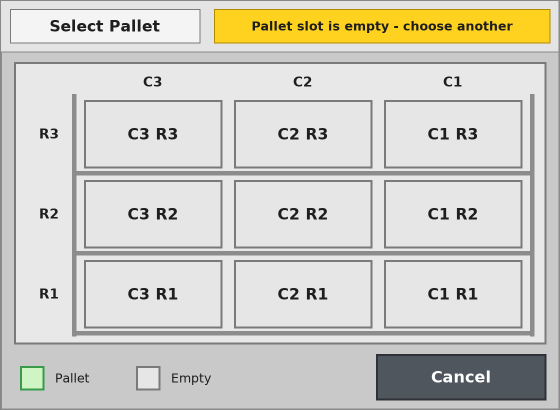
VISUALIZATION SelectPalletDialog  // 560x410
    Rectangle (0,0 560x410)
    Rectangle (0,0 560x52)
    Rectangle (10,9 190x34), "Select Pallet"
    Rectangle (214,12 334x28), "Tap a green slot to retrieve the pallet"
    RoundedRectangle (14,62 532x282)
    Rectangle (84,70 138x24), "C3"
    Rectangle (234,70 138x24), "C2"
    Rectangle (384,70 138x24), "C1"
    Rectangle (24,100 50x68), "R3"
    Rectangle (24,180 50x68), "R2"
    Rectangle (24,260 50x68), "R1"
    Rectangle (72,94 4x242)
    Rectangle (530,94 4x242)
    Rectangle (72,171 462x4)
    Rectangle (72,251 462x4)
    Rectangle (72,331 462x4)
    RoundedRectangle (84,100 138x68), "C3 R3", colour toggle: MAIN.slotOccupied[3,3], invisible if: MAIN.slotEmpty[3,3], input disabled if: MAIN.slotEmpty[3,3]
        OnMouseUp: execute {
            // Only a green box (pallet on the slot) can be chosen
            IF MAIN.slotOccupied[3,3] THEN
                MAIN.selectedColumn := 3;
                MAIN.selectedRow    := 3;
                MAIN.userRequest    := TRUE;
                MAIN.showSlotEmpty  := FALSE;
            END_IF
        }
        OnMouseUp: CloseDialog Dialog=SelectPalletDialog, Result=OK, NumpadKeypadSet=True
    RoundedRectangle (234,100 138x68), "C2 R3", colour toggle: MAIN.slotOccupied[2,3], invisible if: MAIN.slotEmpty[2,3], input disabled if: MAIN.slotEmpty[2,3]
        OnMouseUp: execute {
            // Only a green box (pallet on the slot) can be chosen
            IF MAIN.slotOccupied[2,3] THEN
                MAIN.selectedColumn := 2;
                MAIN.selectedRow    := 3;
                MAIN.userRequest    := TRUE;
                MAIN.showSlotEmpty  := FALSE;
            END_IF
        }
        OnMouseUp: CloseDialog Dialog=SelectPalletDialog, Result=OK, NumpadKeypadSet=True
    RoundedRectangle (384,100 138x68), "C1 R3", colour toggle: MAIN.slotOccupied[1,3], invisible if: MAIN.slotEmpty[1,3], input disabled if: MAIN.slotEmpty[1,3]
        OnMouseUp: execute {
            // Only a green box (pallet on the slot) can be chosen
            IF MAIN.slotOccupied[1,3] THEN
                MAIN.selectedColumn := 1;
                MAIN.selectedRow    := 3;
                MAIN.userRequest    := TRUE;
                MAIN.showSlotEmpty  := FALSE;
            END_IF
        }
        OnMouseUp: CloseDialog Dialog=SelectPalletDialog, Result=OK, NumpadKeypadSet=True
    RoundedRectangle (84,180 138x68), "C3 R2", colour toggle: MAIN.slotOccupied[3,2], invisible if: MAIN.slotEmpty[3,2], input disabled if: MAIN.slotEmpty[3,2]
        OnMouseUp: execute {
            // Only a green box (pallet on the slot) can be chosen
            IF MAIN.slotOccupied[3,2] THEN
                MAIN.selectedColumn := 3;
                MAIN.selectedRow    := 2;
                MAIN.userRequest    := TRUE;
                MAIN.showSlotEmpty  := FALSE;
            END_IF
        }
        OnMouseUp: CloseDialog Dialog=SelectPalletDialog, Result=OK, NumpadKeypadSet=True
    RoundedRectangle (234,180 138x68), "C2 R2", colour toggle: MAIN.slotOccupied[2,2], invisible if: MAIN.slotEmpty[2,2], input disabled if: MAIN.slotEmpty[2,2]
        OnMouseUp: execute {
            // Only a green box (pallet on the slot) can be chosen
            IF MAIN.slotOccupied[2,2] THEN
                MAIN.selectedColumn := 2;
                MAIN.selectedRow    := 2;
                MAIN.userRequest    := TRUE;
                MAIN.showSlotEmpty  := FALSE;
            END_IF
        }
        OnMouseUp: CloseDialog Dialog=SelectPalletDialog, Result=OK, NumpadKeypadSet=True
    RoundedRectangle (384,180 138x68), "C1 R2", colour toggle: MAIN.slotOccupied[1,2], invisible if: MAIN.slotEmpty[1,2], input disabled if: MAIN.slotEmpty[1,2]
        OnMouseUp: execute {
            // Only a green box (pallet on the slot) can be chosen
            IF MAIN.slotOccupied[1,2] THEN
                MAIN.selectedColumn := 1;
                MAIN.selectedRow    := 2;
                MAIN.userRequest    := TRUE;
                MAIN.showSlotEmpty  := FALSE;
            END_IF
        }
        OnMouseUp: CloseDialog Dialog=SelectPalletDialog, Result=OK, NumpadKeypadSet=True
    RoundedRectangle (84,260 138x68), "C3 R1", colour toggle: MAIN.slotOccupied[3,1], invisible if: MAIN.slotEmpty[3,1], input disabled if: MAIN.slotEmpty[3,1]
        OnMouseUp: execute {
            // Only a green box (pallet on the slot) can be chosen
            IF MAIN.slotOccupied[3,1] THEN
                MAIN.selectedColumn := 3;
                MAIN.selectedRow    := 1;
                MAIN.userRequest    := TRUE;
                MAIN.showSlotEmpty  := FALSE;
            END_IF
        }
        OnMouseUp: CloseDialog Dialog=SelectPalletDialog, Result=OK, NumpadKeypadSet=True
    RoundedRectangle (234,260 138x68), "C2 R1", colour toggle: MAIN.slotOccupied[2,1], invisible if: MAIN.slotEmpty[2,1], input disabled if: MAIN.slotEmpty[2,1]
        OnMouseUp: execute {
            // Only a green box (pallet on the slot) can be chosen
            IF MAIN.slotOccupied[2,1] THEN
                MAIN.selectedColumn := 2;
                MAIN.selectedRow    := 1;
                MAIN.userRequest    := TRUE;
                MAIN.showSlotEmpty  := FALSE;
            END_IF
        }
        OnMouseUp: CloseDialog Dialog=SelectPalletDialog, Result=OK, NumpadKeypadSet=True
    RoundedRectangle (384,260 138x68), "C1 R1", colour toggle: MAIN.slotOccupied[1,1], invisible if: MAIN.slotEmpty[1,1], input disabled if: MAIN.slotEmpty[1,1]
        OnMouseUp: execute {
            // Only a green box (pallet on the slot) can be chosen
            IF MAIN.slotOccupied[1,1] THEN
                MAIN.selectedColumn := 1;
                MAIN.selectedRow    := 1;
                MAIN.userRequest    := TRUE;
                MAIN.showSlotEmpty  := FALSE;
            END_IF
        }
        OnMouseUp: CloseDialog Dialog=SelectPalletDialog, Result=OK, NumpadKeypadSet=True
    RoundedRectangle (20,366 24x24)
    Rectangle (52,364 80x28), "Pallet"
    RoundedRectangle (136,366 24x24)
    Rectangle (168,364 80x28), "Empty"
    RoundedRectangle (376,354 170x46), "Cancel"
        OnMouseUp: execute {
            MAIN.cancelRequest := TRUE;   // no pallet chosen: the SFC goes back to Step_10
        }
        OnMouseUp: CloseDialog Dialog=SelectPalletDialog, Result=Cancel, NumpadKeypadSet=True
    RoundedRectangle (384,260 138x68), "C1 R1", colour toggle: MAIN.slotOccupied[1,1], invisible if: MAIN.slotOccupied[1,1], input disabled if: MAIN.slotOccupied[1,1]
        OnMouseUp: execute {
            MAIN.showSlotEmpty := TRUE;   // empty slot: show the message, the dialog stays open
        }
    RoundedRectangle (384,180 138x68), "C1 R2", colour toggle: MAIN.slotOccupied[1,2], invisible if: MAIN.slotOccupied[1,2], input disabled if: MAIN.slotOccupied[1,2]
        OnMouseUp: execute {
            MAIN.showSlotEmpty := TRUE;   // empty slot: show the message, the dialog stays open
        }
    RoundedRectangle (384,100 138x68), "C1 R3", colour toggle: MAIN.slotOccupied[1,3], invisible if: MAIN.slotOccupied[1,3], input disabled if: MAIN.slotOccupied[1,3]
        OnMouseUp: execute {
            MAIN.showSlotEmpty := TRUE;   // empty slot: show the message, the dialog stays open
        }
    RoundedRectangle (234,260 138x68), "C2 R1", colour toggle: MAIN.slotOccupied[2,1], invisible if: MAIN.slotOccupied[2,1], input disabled if: MAIN.slotOccupied[2,1]
        OnMouseUp: execute {
            MAIN.showSlotEmpty := TRUE;   // empty slot: show the message, the dialog stays open
        }
    RoundedRectangle (234,180 138x68), "C2 R2", colour toggle: MAIN.slotOccupied[2,2], invisible if: MAIN.slotOccupied[2,2], input disabled if: MAIN.slotOccupied[2,2]
        OnMouseUp: execute {
            MAIN.showSlotEmpty := TRUE;   // empty slot: show the message, the dialog stays open
        }
    RoundedRectangle (234,100 138x68), "C2 R3", colour toggle: MAIN.slotOccupied[2,3], invisible if: MAIN.slotOccupied[2,3], input disabled if: MAIN.slotOccupied[2,3]
        OnMouseUp: execute {
            MAIN.showSlotEmpty := TRUE;   // empty slot: show the message, the dialog stays open
        }
    RoundedRectangle (84,260 138x68), "C3 R1", colour toggle: MAIN.slotOccupied[3,1], invisible if: MAIN.slotOccupied[3,1], input disabled if: MAIN.slotOccupied[3,1]
        OnMouseUp: execute {
            MAIN.showSlotEmpty := TRUE;   // empty slot: show the message, the dialog stays open
        }
    RoundedRectangle (84,180 138x68), "C3 R2", colour toggle: MAIN.slotOccupied[3,2], invisible if: MAIN.slotOccupied[3,2], input disabled if: MAIN.slotOccupied[3,2]
        OnMouseUp: execute {
            MAIN.showSlotEmpty := TRUE;   // empty slot: show the message, the dialog stays open
        }
    RoundedRectangle (84,100 138x68), "C3 R3", colour toggle: MAIN.slotOccupied[3,3], invisible if: MAIN.slotOccupied[3,3], input disabled if: MAIN.slotOccupied[3,3]
        OnMouseUp: execute {
            MAIN.showSlotEmpty := TRUE;   // empty slot: show the message, the dialog stays open
        }
    Rectangle (214,9 336x34), "Pallet slot is empty - choose another", invisible if: MAIN.hideSlotEmpty, input disabled if: MAIN.hideSlotEmpty
END_VISUALIZATION

(* stored: Version 1.1.0.1, ProductVersion 3.1.4024.12
   Visu SelectPalletDialog: Id {61ea3e01-3f21-44f3-84fc-9478cd6e9d3c} *)
